PROGRAM MAIN
VAR CONSTANT	
	Axis_Count : INT := 4 ;
END_VAR
VAR
	power : BOOL;
	Index : INT := 1;
	
	AxisList : ARRAY[1..Axis_Count] OF AXIS_REF;
	
	Axis_State:  ARRAY[1..Axis_Count] OF INT;
	Axis_Power : ARRAY[1..Axis_Count] OF MC_Power;
	Axis_Reset : ARRAY[1..Axis_Count] OF MC_Reset;
	Axis_Home : ARRAY[1..Axis_Count] OF MC_Home;
	Axis_MoveAbs : ARRAY[1..Axis_Count] OF ARRAY[0..1] OF MC_MoveAbsolute;
	Axis_ErrorID : ARRAY[1..Axis_Count] OF UDINT;
	absSwitch : ARRAY[1..Axis_Count] OF INT;
	
	bHomeSwitch : ARRAY[1..Axis_Count] OF BOOL;
	startMove : ARRAY[1..Axis_Count] OF BOOL;
	homeBusy : ARRAY[1..Axis_Count] OF BOOL; // check if home function block is busy
	actPos : ARRAY[1..Axis_Count] OF LREAL; // array of actual position of each axis
	
	Axis_GoalPos : LREAL;
	
	rMoveVelocity : LREAL := 1600;//42666;
	rMoveAcceleration : LREAL := 12000;//120000;
	rMoveDecceleration : LREAL := 12000;//120000;
	rMoveJerk : LREAL := 560000;
	
	iCycleNum : DINT := 0;
END_VAR

iCycleNum := iCycleNum + 1;
FOR Index := 1 TO Axis_Count BY 1 DO
	AxisList[Index].ReadStatus();
	Axis_Power[Index](Axis:=AxisList[Index], Enable:=power, Enable_Positive:=TRUE, Enable_Negative:=TRUE);
	IF power THEN
		homeBusy[Index] := Axis_Home[Index].Busy;
		actPos[Index] := AxisList[Index].NcToPlc.ActPos;
		Axis_MoveAbs[Index][0](Axis:=AxisList[Index], Execute:=FALSE);
		Axis_MoveAbs[Index][1](Axis:=AxisList[Index], Execute:=FALSE);
		CASE Axis_State[Index] OF
			0: // Initial
				Axis_Reset[Index](Axis:=AxisList[Index], Execute := FALSE);
				absSwitch[Index] := 0;
				Axis_State[Index] := 10;
			10: // Start Drive Reset
				Axis_Reset[Index](Axis:=AxisList[Index], Execute := TRUE); 
				IF Axis_Reset[Index].Done THEN
					Axis_State[Index] := 20;
				ELSIF Axis_Reset[Index].Error THEN
					Axis_ErrorID[Index] := Axis_Reset[Index].ErrorID;
					Axis_State[Index] := 997;
				END_IF
			20: // Wait for Drive to Reset
				IF Axis_Power[Index].Status THEN
					Axis_State[Index] := 30;
				//ELSE
				//	Axis_State[Index] := 996;
				//	Axis_ErrorID[Index] := Axis_Power[Index].ErrorID;
				END_IF
			30: // Set current position / Homing
				IF bHomeSwitch[Index] THEN
					Axis_Home[Index](Axis:=AxisList[Index], HomingMode:=MC_HomingMode.MC_Direct, Position:=Axis_GoalPos, Execute:=TRUE);
					IF Axis_Home[Index].Error THEN
						Axis_State[Index] := 998;
					END_IF
					IF Axis_Home[Index].Done THEN
						Axis_Home[Index](Axis:=AxisList[Index], Execute:=FALSE);
						bHomeSwitch[Index] := FALSE;
					END_IF 
				ELSIF startMove[Index] THEN
					startMove[Index] := FALSE;
					Axis_State[Index] := 40;
				END_IF
			40: // Start Absolute Move
				IF Axis_MoveAbs[Index][absSwitch[Index]].Busy THEN
					absSwitch[Index] := (absSwitch[Index] + 1) MOD 2;
				END_IF
				Axis_MoveAbs[Index][absSwitch[Index]](Axis:=AxisList[Index], Position := Axis_GoalPos, BufferMode := MC_Aborting, Velocity := rMoveVelocity,
							Acceleration := rMoveAcceleration, Deceleration := rMoveDecceleration, Jerk := rMoveJerk, Execute := TRUE);
				IF Axis_MoveAbs[Index][absSwitch[Index]].Error THEN //Axis_MoveAbs.Done AND 
					Axis_State[Index] := 999;
				END_IF
				Axis_State[Index] := 30;
			
			999: //Error Fixing (TODO)
		END_CASE
	END_IF
END_FOR

END_PROGRAM

(* stored: Version 1.1.0.1, ProductVersion 3.1.4024.9
   POU MAIN: Id {31b0bc00-96e9-4e64-af9b-c5575f64f6fc}, SpecialFunc None *)
